// TIA Portal V21 export
// export: Created 2026-11-10T19:16:33.612469Z, ExportSetting WithDefaults, DisplayName Totally Integrated Automation Portal, DisplayVersion V21 Update 3, DisplayName STEP 7 Professional, DisplayVersion V21 Update 3, DisplayName STEP 7 Safety, DisplayVersion V21, DisplayName Tech WebApplication, DisplayVersion V21, DisplayName WinCC Basic/Comfort/Advanced, DisplayVersion V21 Update 3, DisplayName WinCC Unified, DisplayVersion V21 Update 3
TYPE "UDT_300"
// stored: IsFailsafeCompliant false
   STRUCT
      "a" : Int := 3;
      "b" : Real;
      c : Array[0..1] of Bool;
   END_STRUCT;
END_TYPE
